Yaskawa INFORM job: CLEAN_R1.JBI

/JOB
//NAME CLEAN_R1
//POS
///NPOS 12,0,0,3,0,0
///TOOL 0
///POSTYPE PULSE
///PULSE
C00000=-109209,-54646,-76367,1352,-34711,-1501
C00001=-109209,-55063,-81056,1461,-31794,-1563
C00002=-109209,-55028,-89231,1746,-26136,-1717
C00003=-109209,-54990,-79963,1432,-32492,-1548
C00004=-125064,-56796,-80702,-11384,-34301,7100
C00005=-125064,-57070,-84860,-12217,-31699,7569
C00006=-125064,-56546,-78346,-10989,-35705,6872
C00007=-107494,-54447,-77481,2777,-33833,-2456
C00008=-111906,-43067,-86202,-1367,-19196,245
C00009=-112783,-41007,-86214,-2792,-17657,1092
C00010=-111636,-45955,-87712,-948,-20329,-5
C00011=-111636,-46808,-68835,-590,-33981,-193
P00001=-112783,-40998,-86242,-2796,-17631,1094
P00100=0,-60000,-60000,0,-90000,0
P00101=-130000,-60000,-60000,0,-90000,0
//INST
///DATE 2025/07/15 15:21
///ATTR SC,RW
///GROUP1 RB1
///LVARS 0,1,0,0,0,0,0,0
NOP
SET LI000 100
MOVJ P100 VJ=50.00
MOVJ P101 VJ=50.00
MOVJ C00000 VJ=50.00
MOVJ C00001 VJ=50.00
WAIT IN#(12)=ON
MOVL C00002 V=750.0 PL=0
PULSE OT#(9) T=1.00
PULSE OT#(10) T=1.00
TIMER T=2.00
WAIT IN#(12)=ON
TIMER T=0.20
MOVL C00003 V=750.0 PL=0
MOVL C00004 V=750.0 PL=0
MOVL C00005 V=750.0 PL=0
PULSE OT#(11) T=0.30
TIMER T=0.60
MOVL C00006 V=750.0 PL=0
MOVL C00007 V=750.0 PL=0
MOVL C00008 V=750.0
PULSE OT#(4095) T=0.75
TIMER T=1.00
MOVL C00009 V=750.0 PL=0
MOVL P001 V=23.0
TIMER T=0.25
PULSE OT#(12) T=0.50
TIMER T=0.50
MOVL C00010 V=750.0
MOVL C00011 V=750.0
MOVJ P101 VJ=50.00
MOVJ P100 VJ=50.00
SET I097 0
END
